Fanuc KAREL source: kt00414.KL

-- PROVISIONAL review KL for V770-1; original PC SHA256 fbbd6e2345d7589313c7fea6683c9997bc40f32f276ed45ecbf103da14ea998f
-- Incomplete behavior may be omitted. Consult companion uncertainty JSON. Do not deploy.
PROGRAM KT00414
%NOLOCKGROUP
VAR
  OUT : BOOLEAN
-- UNRESOLVED_DECL Y1 type=002018
-- UNRESOLVED_DECL H2 type=002017
BEGIN
  -- UNRESOLVED_PC offsets 5-19; opcodes 2E,22,9D,33,B2
  -- UNRESOLVED_PC offsets 24-38; opcodes 2E,22,9D,33,B4
  -- UNRESOLVED_PC offsets 43-68; opcodes 22,9D,33,B1,22,9D,33,B3,5B,23
  -- UNRESOLVED_PC offsets 73-77; opcodes 7F
END KT00414
